// TIA Portal V20 export
Screen "Pop-up_SYSTEM_RTSTOP_Popup"  210x126
  ScreenItem "Background" at 0,0 size 210x126  Type=HmiRectangle
  ScreenItem "Descr_SafateyDialog" at 2,26 size 180x25  Type=HmiTextBox
  ScreenItem "Overview_SafetyDialog" at 1,1 size 208x25  Type=HmiTextBox
  ScreenItem "Cancel Mode" at 110,56 size 90x60  Type=HmiButton
  ScreenItem "Stop_RT" at 10,56 size 90x60  Type=HmiButton
